Fanuc KAREL source: KD00026.KL

PROGRAM KD00026
%NOLOCKGROUP
VAR
  I: INTEGER
  J: INTEGER
  B: BOOLEAN
  R: REAL
  S: STRING[80]
BEGIN
  CONDITION[1]:
  WHEN DIN[1] = ON DO
    I = 1
  ENDCONDITION
END KD00026
